ADAPTER arm (* Adapter Interface *)
  (* Standard: 61499-1 *)
  (* Version 0.0, 10/22/2026, lizar, Schneider Electric *)
  PACKAGE Main;
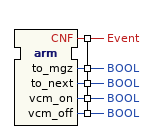
  EVENT_OUTPUT
    CNF WITH to_mgz, to_next, vcm_on, vcm_off; (* Confirmation from Plug *)
  END_EVENT
  VAR_OUTPUT
    to_mgz : BOOL; (* Indication Data from Plug *)
    to_next : BOOL; (* Indication Data from Plug *)
    vcm_on : BOOL; (* Indication Data from Plug *)
    vcm_off : BOOL; (* Indication Data from Plug *)
  END_VAR
  SERVICE SOCKET/PLUG
    SEQUENCE request_confirm
      SOCKET.REQ(REQD) -> PLUG.REQ(REQD);
      PLUG.CNF(CNFD) -> SOCKET.CNF(CNFD);
    END_SEQUENCE
    SEQUENCE indication_response
      PLUG.IND(to_mgz) -> SOCKET.IND(to_mgz);
      SOCKET.RSP(RSPD) -> PLUG.RSP(RSPD);
    END_SEQUENCE
  END_SERVICE
END_ADAPTER
